// TIA Portal V20 export
// export: Created 2026-10-12T05:42:28.8738101Z, ExportSetting WithDefaults, DisplayName Totally Integrated Automation Portal, DisplayVersion V20, DisplayName TIA Portal Openness, DisplayVersion V20, DisplayName TIA Portal Teamcenter Gateway, DisplayVersion V20, DisplayName TIA Portal Version Control Interface, DisplayVersion V20, DisplayName SINAMICS Startdrive Advanced, DisplayVersion V20 SP1 Update 2, DisplayName SINAMICS Startdrive G110M, G120, G120C, G120D, G120P, G115D, DisplayVersion V20 SP1 Update 2, DisplayName SINAMICS Startdrive G130, G150, S120, S150, SINAMICS MV, G220, S200, S210, DisplayVersion V20 SP1 Update 2, DisplayName STEP 7 Professional, DisplayVersion V20, DisplayName STEP 7 Safety, DisplayVersion V20, DisplayName WinCC Basic/Comfort/Advanced, DisplayVersion V20, DisplayName WinCC Professional, DisplayVersion V20, DisplayName WinCC Unified, DisplayVersion V20
FUNCTION "FRK_ConfigBegin" : Void   // FC23, SCL
{ S7_Optimized_Access := 'TRUE' }
VERSION : 0.1
// stored: AutoNumber true, IsIECCheckEnabled false, SetENOAutomatically false, UDAEnableTagReadback false
   VAR_INPUT
      PageIndex : DInt;
      Revision : UDInt;
   END_VAR
   VAR_IN_OUT
      Cursor : "FRK_ConfigCursor";
      Page : "ST_ConfigPage";
   END_VAR
   VAR_TEMP
      Index : Int;
   END_VAR
BEGIN

   #Cursor.Position := 0;
   #Cursor.First := 0;
   #Page.Revision := #Revision;
   #Page.PageIndex := 0;
   IF #PageIndex >= 0 AND #PageIndex <= 32767 THEN
       #Cursor.First := #PageIndex * 16;
       #Page.PageIndex := DINT_TO_INT(#PageIndex);
   END_IF;
   #Page.PageCount := 1;
   #Page.EntryCount := 0;
   "FRK_UnitScratch".EmptyConfigEntry.ValueType := 1;
   "FRK_UnitScratch".EmptyConfigEntry.Readable := TRUE;
   FOR #Index := 1 TO 16 DO
       #Page.Entries[#Index] := "FRK_UnitScratch".EmptyConfigEntry;
   END_FOR;
END_FUNCTION
